// System API/SEC/API/bds_sec_saveSecret
/// This API function is used to store a 16 byte secret key for a specific security access level.
///
///=======
/// Remarks:
///=======
///
///   + The secret keys are stored in an encrypted flash section of the Hardware Security Module (HSM) and cannot be read out.
///   + This asynchronous function must be called several times until the result is available.
///   + If there is no HSM access conflict with another instance, the completion of this function (execution within a loop) takes
///	   + about 1250us (microseconds) with a new secret key and
///	   + about 350us (microseconds) with the same secret key as already stored.
///   + This function will be rejected if another asynchronous security function was already started for this instance.
///
///----------
/// FFI:
///----------
///This API can be used in trusted partitions only. See Freedom from Interference (FFI) concept for more details.
///
///----------
/// Attention:
///----------
///
///   + This function writes the secret key physically into the HSM flash. Therefore this function should not be called cyclically.
///   + Do not interrupt this function by power off to prevent corrupted secret keys.
///
///==================================================================		  			===================================================================================================
///Return value    								  									Description
///==================================================================		  			===================================================================================================
///16#0000: BDS_SEC_ERR_NO_ERROR_DU16													Function was executed without errors. The provided secret key was stored in HSM.
///16#0001: BDS_SEC_ERR_PARAM1_ERROR_DU16												Invalid instance number. 
///16#0002: BDS_SEC_ERR_PARAM2_ERROR_DU16												Invalid access level.
///16#0003: BDS_SEC_ERR_PARAM3_ERROR_DU16												Invalid secret key pointer. Pointer is equal to zero.
///16#0010: BDS_SEC_ERR_REQUEST_PENDING_DU16											This asynchronous function was not yet completed and must be called again with the same parameter values. Several function calls may be required in particular if another security manager instance is also running.
///16#0020:BDS_SEC_ERR_INVALID_SEQUENCE_DU16											This function was called although another asynchronous security function was not yet completed. The other asynchronous function that has already been started must be called again and must be completed before this function can be started.
///16#0033: BDS_SEC_ERR_OPEN_SESSION_FAILED_DU16										Security session could not be opened for this function.Possible reason could be that the HSM is not running. 
///16#0035: BDS_SEC_ERR_CLOSE_SESSION_FAILED_DU16										Security session could not be closed for this function. 
///16#0038: BDS_SEC_ERR_SET_PASSWORD_FAILED_DU16										The internal storage of the secret key failed. To terminate the function, it must be called again.
///
///==================================================================		   			===================================================================================================
///
///For Access levels, Refer the below table & provide the value,
///
///==================================================================		  			===================================================================================================
///Access Level Variable   								  							Value
///==================================================================		  			===================================================================================================
///BDS_SEC_ACC_LEVEL_0_E																0
///BDS_SEC_ACC_LEVEL_1_E																1
///BDS_SEC_ACC_LEVEL_2_E																2
///BDS_SEC_ACC_LEVEL_3_E																3
///BDS_SEC_ACC_LEVEL_4_E																4
///BDS_SEC_ACC_LEVEL_5_E																5
///BDS_SEC_ACC_LEVEL_6_E																6
///BDS_SEC_ACC_LEVEL_7_E																7
///BDS_SEC_ACC_LEVEL_8_E																8
///BDS_SEC_ACC_LEVEL_9_E																9
///BDS_SEC_ACC_LEVEL_10_E																10
///BDS_SEC_ACC_LEVEL_11_E																11
///BDS_SEC_ACC_LEVEL_12_E																12
///BDS_SEC_ACC_LEVEL_13_E																13
///BDS_SEC_ACC_LEVEL_14_E																14
///BDS_SEC_ACC_LEVEL_15_E																15
///BDS_SEC_ACC_LEVEL_16_E																16
///BDS_SEC_ACC_LEVEL_17_E																17
///BDS_SEC_ACC_LEVEL_18_E																18
///BDS_SEC_ACC_LEVEL_19_E																19
///BDS_SEC_ACC_LEVEL_20_E																20
///
///==================================================================		   			===================================================================================================
///
///=======
///Code Example:
///=======
///============================================================================
///
///PROGRAM appl_Task_1
///
///  VAR
///	return_u16 : UINT;
///
///	secKey_au8 : STRING(16);
///	
///  END_VAR
///  
///  (*check for request to store a new secret key*)
///
/// secKey_au8 :=  'MyNewKey' 
///
///result_u16 := bds_sec_saveSecret(bds_diag_inst_te.BDS_SEC_ASW_INST_NAME_1_E, 1, ADR(secKey_au8));
///
///============================================================================
///
{attribute 'external_name' := 'cmp_rts_bds_sec_saveSecret'}
FUNCTION bds_sec_saveSecret : UINT
VAR_INPUT
	///Instance number. pointer to |bds_diag_inst_te|
	diagInst_e: bds_diag_inst_te;
	///Pointer to a variable which must be provided(Refer access level table). The current level will be copied to this variable. 
	level_e: USINT;
	///Pointer to a 16 byte buffer which must be provided by the application and which must contain the new secret key.
	secrKey_pau8: POINTER TO USINT;
END_VAR

END_FUNCTION

// System API/SEC/API/bds_sec_scrambleRexrothSecretsPerm
///This API function is used to scramble all internally stored Rexroth secret keys.
///
///=======
/// Remarks:
///=======
///
///   + This asynchronous function must be called several times until the final result is available.
///   + The completion of this function (execution within a loop) takes about 5,3ms if there is no HSM access conflict with another instance.
///   + This function will be rejected if another asynchronous security function was already started for this instance.
///
///----------
/// FFI:
///----------
///This API can be used in trusted partitions only. See Freedom from Interference (FFI) concept for more details.
///
///----------
/// Attention:
///----------
///
///This function cannot be undone! After the execution of this function the corresponding Rexroth access levels can not be activated any more. This excludes Rexroth personnel from diagnosis information that might be required in case of field service or field claims irrevocably. 
///   
///----------
/// Info:
///----------
///
///This function writes the secret keys physically into the HSM flash. Therefore this function should not be called cyclically.
///   
///==================================================================		  			===================================================================================================
///Return value    								  									Description
///==================================================================		  			===================================================================================================
///16#0000: BDS_SEC_ERR_NO_ERROR_DU16													Function was executed without errors
///16#0010: BDS_SEC_ERR_REQUEST_PENDING_DU16											This asynchronous function was not yet completed and must be called again with the same parameter values. Several function calls may be required in particular if another security manager instance is also running.
///16#0020: BDS_SEC_ERR_INVALID_SEQUENCE_DU16											This function was called although another asynchronous security function was not yet completed. The other asynchronous function that has already been started must be called again and must be completed before this function can be started.
///16#0033: BDS_SEC_ERR_OPEN_SESSION_FAILED_DU16										Security session could not be opened for this function.Possible reason could be that the HSM is not running. 
///16#0034: BDS_SEC_ERR_GENERATE_RANDOM_FAILED_DU16										The process to generate the random has been failed.  To terminate the function, it must be called again.
///16#0035: BDS_SEC_ERR_CLOSE_SESSION_FAILED_DU16										Security session could not be closed for this function. 
///16#0038: BDS_SEC_ERR_SET_PASSWORD_FAILED_DU16										The internal storage of the secret key failed. To terminate the function, it must be called again.
///
///==================================================================		   			===================================================================================================
///
///
///=======
///Code Example:
///=======
///============================================================================
///
///PROGRAM appl_Task_1
///
///  VAR
///	
///  END_VAR
///  
///  (*check if Rexroth access levels shall be scrambled & call the API*)
///  
///result_u16 := bds_sec_scrambleRexrothSecretsPerm();
///
///============================================================================
///
{attribute 'external_name' := 'cmp_rts_bds_sec_scrambleRexrothSecretsPerm'}
FUNCTION bds_sec_scrambleRexrothSecretsPerm : UINT

END_FUNCTION

// System API/SYS/API/bds_sys_ait
///This function gets the temperature of the printed circuit board (PCB)
///
///=======
/// Remarks:
///=======
///    + The voltage of the NTC thermistor located on the PCB is transferred into temperature between -40..150°C.
///    + The resolution is 1°C .
///    + The |GVL_sys| is given for usage of defines.
///    + Import the bds_rts_ec.xml to use the enums. (Refer example below).
///
///----------
/// FFI:
///----------
///This API can be used in trusted partitions only. See Freedom from Interference (FFI) concept for more details.
///
///==================================================================		  			===================================================================================================
///Return value    								  									Description
///==================================================================		  			===================================================================================================
///16#00																				No error.
///16#01																				A parameter is invalid.
///16#02																				Function call was erroneous.
///
///==================================================================		   			===================================================================================================
///
///=======
///Code Example:
///=======
///============================================================================
///
///PROGRAM appl_10ms_task
///
///VAR
///	tsg1_value_s16: INT := 16#00;
///END_VAR
///
///(* get a temperature 1 of high temperature of hardware*)
///
///bds_sys_ait(bds_sys_ait_signal_te.TSGI1, ADR(tsg1_value_s16));
///
///============================================================================
{attribute 'external_name' := 'cmp_rts_bds_sys_ait'}
FUNCTION bds_sys_ait : USINT
VAR_INPUT
	///The assigned signal name of the input.
	signal_e: UINT;
	///Storage address of the value.
	///
	///Range:
	///-40..150 [°C]
	value_ps16: POINTER TO INT;
END_VAR

END_FUNCTION

// System API/SYS/API/bds_sys_aiv
///This function gets the voltage of the analog system input.
///
///=======
/// Remarks:
///=======
///    + Enable the access to all system voltages [mV].
///    + The |GVL_sys| is given for usage of defines.
///    + Import the bds_rts_ec.xml to use the enums. (Refer example below).
///
///----------
/// FFI:
///----------
///This API can be used in trusted partitions only. See Freedom from Interference (FFI) concept for more details.
///	
///==================================================================		  			===================================================================================================
///Return value    								  									Description
///==================================================================		  			===================================================================================================
///16#00																				No error.
///16#01																				A parameter is invalid.
///16#02																				Function call was erroneous.
///
///==================================================================		   			===================================================================================================
///
///=======
///Code Example:
///=======
///============================================================================
///
///PROGRAM appl_10ms_task
///
///VAR
///
///	state_VSS4_u16: UINT := 16#00;
///
///END_VAR
///
///
///(* get a sensor supply voltage *)
///
///bds_sys_aiv(bds_sys_aiv_signal_te.VSS4V10, ADR(state_VSS4_u16));
///
///
///============================================================================
{attribute 'external_name' := 'cmp_rts_bds_sys_aiv'}
FUNCTION bds_sys_aiv : USINT
VAR_INPUT
	///The signal name of the input.
	signal_e: UINT;
	///Storage address of the value.
	///
	///Range:
	///0..40000 [mV]
	value_pu16: POINTER TO UINT;
END_VAR

END_FUNCTION

// System API/SYS/API/bds_sys_cancelAltWakeup
///This function transitions the ECU operating state from RUN to POSTRUN, when the system wakeup reason is not T15. For different methods of ECU wakeup mechanisms please refer page Wakeup.
///
///=======
/// Remarks:
///=======
///    + This function has to be called when the ECU is in RUN state. 
///    + This is most suitable for applications where T15 is not used to switch the ECU OFF.
///    + Wakeup source information can be identified using the BSW API |bds_sys_getResetInfo|.
///    + BSW API |bds_sys_releasePostRunProlong| is used to transition the ECU operating state from POSTRUN to SHUTDOWN.
///    + The |GVL_sys| is given for usage of defines.
///	
///----------
/// FFI:
///----------
///This API can be used in trusted partitions only. See Freedom from Interference (FFI) concept for more details.
///
///----------
/// NOTICE:
///----------
///    + This function has no effect when ECU wakeup has occurred by T15.
///	
///==================================================================		  			===================================================================================================
///Return value    								  									Description
///==================================================================		  			===================================================================================================
///0																					ECU Operating state has moved from RUN to POSTRUN.
///1																					T15 (Ignition pin) is ON.x
///																					    + Note: This return value appears also when ECU woke up by CAN and then T15 turns ON, before this function is called. So, after this, to transition the ECU to POSTRUN state T15 should be turned OFF.
///2																					ECU is already in POSTRUN state.
///
///==================================================================		   			===================================================================================================
///
///=======
///Code Example:
///=======
///============================================================================
///
///PROGRAM PRG
///
///VAR
///
///	return_u8 : USINT;
///
/// flag_u8 :USINT;
///
///END_VAR
///
///IF(0 = flag_u8) THEN
///
/// bds_sys_requestPostRunProlong(); (* request for prolong in POSTRUN*)
///
///	return_u8 := bds_sys_cancelAltWakeup(); (*forces system state to go to POSTRUN*)
///
/// bds_sys_releasePostrunProlong(); (*transitions system state from POSTRUN to SHUTDOWN*)
///
/// flag_u8:=1;
///
///END_IF
///
///============================================================================
{attribute 'external_name' := 'cmp_rts_bds_sys_cancelAltWakeup'}
FUNCTION bds_sys_cancelAltWakeup : USINT

END_FUNCTION

// System API/SYS/API/bds_sys_getResetInfo
///This function can be used in order to get information about reset of ECU.
///
///=======
/// Remarks:
///=======
///    + This function should be used in case of reset problems. The Rexroth service needs this info for solving the problem.
///    + The reset information will only be cleared after power on.
///    + The Reset IDs & Reset Group IDs can be found in "rba_Reset_Cfg.h" header file. All the Reset group IDs are listed down under enum variable "rba_Reset_Grp_ten" and all the reset IDs are listed down under enum variable "rba_Reset_Id_ten".
///    + The |GVL_sys| is given for usage of defines.
///
///----------
/// FFI:
///----------
///This API can be used in trusted partitions . For untrusted partitions use |bds_sys_getResetInfo_ffi|. See Freedom from Interference (FFI) concept for more details.
///
///==================================================================		  			===================================================================================================
///Return value    								  									Description
///==================================================================		  			===================================================================================================
///16#0000																				No error. 
///16#0001																				Function called with null pointer.
///16#25																				FFI API access error.
///
///==================================================================		   			===================================================================================================
///=======
///Code Example:
///=======
///============================================================================
///
///PROGRAM appl_10ms_task
///
///VAR
///
///	reset_info : bds_ResetInfo_ts;
///	
///	return_u8 : UINT;
///
///END_VAR
///
///return_u8 := bds_sys_getResetInfo(ADR(reset_info)); (*reads the reset information of ECU*)
///
///============================================================================
{attribute 'external_name' := 'cmp_rts_bds_sys_getResetInfo'}
FUNCTION bds_sys_getResetInfo : UINT
VAR_INPUT
	///Pointer to |bds_ResetInfo_ts|
	resetinfo_ps: POINTER TO bds_ResetInfo_ts;
END_VAR

END_FUNCTION

// System API/SYS/FFI_API/bds_sys_getResetInfo_ffi
{attribute 'external_name' := 'cmp_rts_bds_sys_getResetInfo_ffi'}
FUNCTION bds_sys_getResetInfo_ffi : UINT
VAR_INPUT
	///Pointer to |bds_ResetInfo_ts|
	resetinfo_ps: POINTER TO bds_ResetInfo_ts;
END_VAR

END_FUNCTION

// System API/SYS/API/bds_sys_releasePostRunProlong
///This function terminates prolonging of  POSTRUN state and enters to SHUTDOWN state.     
///=======
/// Remarks:
///=======
///    + By calling this function, POSTRUN is terminated, if system is in POSTRUN state and enters to SHUTDOWN phase. 
///    + After calling |bds_sys_requestPostRunProlong| and after completion of tasks in POSTRUN this function must be called. If not, exit from POSTRUN is only through timeout.
///    + The |GVL_sys| is given for usage of defines.
///	
///----------
/// FFI:
///----------
///This API can be used in trusted partitions only. See Freedom from Interference (FFI) concept for more details.
///
///==================================================================		  			===================================================================================================
///Return value    								  									Description
///==================================================================		  			===================================================================================================
///None																				None
///
///==================================================================		   			===================================================================================================
///
///
///=======
///Code Example:
///=======
///============================================================================
///
///PROGRAM appl_1ms_task
///
///VAR
///
///END_VAR
///
///bds_sys_releasePostRunProlong();  (* release of prolong in postrun *)
///
///============================================================================
{attribute 'external_name' := 'cmp_rts_bds_sys_releasePostRunProlong'}
FUNCTION bds_sys_releasePostRunProlong : BOOL

END_FUNCTION

// System API/SYS/API/bds_sys_requestPostRunProlong
///This function enables a prolonging cyclic tasks in POSTRUN.    
///=======
/// Remarks:
///=======
///    + This function can be called in initialization or RUN state of system.
///    + After calling this function, termination from POSTRUN state is possible only by calling |bds_sys_releasePostRunProlong| or Timeout set for POSTRUN prolong.  
///    + The Maximum Post Run timeout allowed is 24hours / 86400 sec. The actual Post Run timeout is configured in easyConfig.In order to shorten the Post Run timeout  the  API |bds_sys_releasePostRunProlong| shall be used.
///    + Without calling this function, No cyclic tasks are in POSTRUN. Only shutdown functions will be executed after Ignition(T15) goes OFF.
///    + The |GVL_sys| is given for usage of defines.
///	
///----------
/// FFI:
///----------
///This API can be used in trusted partitions only. See Freedom from Interference (FFI) concept for more details.
///
///---------
///  NOTICE:
///---------
///Don't forget to call  |bds_sys_releasePostRunProlong|, after enabling cyclic tasks POSTRUN.
///	
///==================================================================		  			===================================================================================================
///Return value    								  									Description
///==================================================================		  			===================================================================================================
///None																				None
///
///==================================================================		   			===================================================================================================
///
///
///=======
///Code Example:
///=======
///============================================================================
///
///PROGRAM appl_1ms_task
///
///VAR
///
///END_VAR
///
///bds_sys_requestPostRunProlong();  (* request for prolong in postrun *)
///
///============================================================================
{attribute 'external_name' := 'cmp_rts_bds_sys_requestPostRunProlong'}
FUNCTION bds_sys_requestPostRunProlong : BOOL

END_FUNCTION

// System API/SYS/API/bds_sys_di
///This function gets the state of a digital system input.
///
///=======
/// Remarks:
///=======
///    + Enable the access to all digital signals.
///    + The |GVL_sys| is given for usage of defines.
///    + Import the bds_rts_ec.xml to use the enums. (Refer example below).
///
///----------
/// FFI:
///----------
///This API can be used in trusted partitions only. See Freedom from Interference (FFI) concept for more details.
///
///==================================================================		  			===================================================================================================
///Return value    								  									Description
///==================================================================		  			===================================================================================================
///16#00																				No error.
///16#01																				A parameter is invalid.
///16#02																				Function call was erroneous.
///
///==================================================================		   			===================================================================================================
///
///=======
///Code Example:
///=======
///============================================================================
///
///PROGRAM appl_10ms_task
///
///VAR
///
///	state_u8: USINT := 16#00;
///
///END_VAR
///
///(* get a state of the inhibit signal *)
///
///bds_sys_di(bds_sys_di_signal_te.ST_INH, ADR(state_u8));
///
///============================================================================
{attribute 'external_name' := 'cmp_rts_bds_sys_di'}
FUNCTION bds_sys_di : USINT
VAR_INPUT
	///The assigned signal name of the input.
	signal_e: UINT;
	///Storage address of the state.
	///
	///States:
	///    + 0 : OFF
	///    + 1 : ON
	state_pu8: POINTER TO USINT;
END_VAR

END_FUNCTION

// System API/SYS/API/bds_sys_getAge
///This function reads the operating time counter of the ECU in minutes.
///
///=======
/// Remarks:
///=======
///    + The counter is incremented by 1 for each minute and saved in non-volatile memory for every 30 minutes.
///    + The operating time counter cannot be reset.
///    + The operating time counter records the total operating time of the device in minutes.
///    + The system time of controller since last reset can be determined using the functions |bds_sys_getTime|.
///    + The |GVL_sys| is given for usage of defines.
///	
///----------
/// FFI:
///----------
///This API can be used in trusted partitions . For untrusted partitions use |bds_sys_getAge_ffi|. See Freedom from Interference (FFI) concept for more details.
///
///----------
/// NOTICE:
///----------
///    + Operating time is saved in case of ignition off event
///    + Operation time is not saved, if ECU power supply is switched off .
///
///==================================================================		  			===================================================================================================
///Return value    								  									Description
///==================================================================		  			===================================================================================================
///Value																				Total operating time of the ECU in minutes
///16#00: BDS_SYS_FFI_ACCESS_ERROR_GETVALUE_DU32										FFI API access error.
///
///==================================================================		   			===================================================================================================
///
///=======
///Code Example:
///=======
///============================================================================
///
///PROGRAM appl_10ms_task
///
///VAR
///
///	operating_hours_u32: UDINT := 16#00;
///
///END_VAR
///
///operating_hours_u32 := bds_sys_getAge(); (* returns Total operating hours of the ECU in minutes *)
///
///============================================================================
{attribute 'external_name' := 'cmp_rts_bds_sys_getAge'}
FUNCTION bds_sys_getAge : UDINT

END_FUNCTION

// System API/SYS/API/bds_sys_getTime
///This function reads the system time of controller since last reset.
///=======
/// Remarks:
///=======
///    + The system time starts at 0 again every time the system is switched on. 
///    + Return value is 64 bit value (counter width).
///    + In order to detect a counter overrun, for long operating times, the operating time counter must also be evaluated using the function |bds_sys_getAge|. 
///    + The |GVL_sys| is given for usage of defines.
///
///----------
/// FFI:
///----------
///This API can be used in trusted partitions . For untrusted partitions use |bds_sys_getTime_ffi|. See Freedom from Interference (FFI) concept for more details.
///
///==================================================================		  			===================================================================================================
///Return value    								  									Description
///==================================================================		  			===================================================================================================
///Value																				System time in microseconds [us].
///16#00: BDS_SYS_FFI_ACCESS_ERROR_GETVALUE_DU64										FFI API access error.
///
///==================================================================		   			===================================================================================================
///
///
///=======
///Code Example:
///=======
///============================================================================
///
///PROGRAM appl_10ms_task
///
///VAR
///
///	operating_time : ULINT := 16#00;
///
///END_VAR
///
///operating_time := bds_sys_getTime();  (* returns Operating time in microseconds since last reset *)
///
///============================================================================
{attribute 'external_name' := 'cmp_rts_bds_sys_getTime'}
FUNCTION bds_sys_getTime : ULINT

END_FUNCTION

// System API/SYS/FFI_API/bds_sys_getTime_ffi
{attribute 'external_name' := 'cmp_rts_bds_sys_getTime_ffi'}
FUNCTION bds_sys_getTime_ffi : ULINT

END_FUNCTION

// System API/SYS/FFI_API/bds_sys_getAge_ffi
{attribute 'external_name' := 'cmp_rts_bds_sys_getAge_ffi'}
FUNCTION bds_sys_getAge_ffi : UDINT

END_FUNCTION

// System API/SYS/API/bds_sys_getCoreLoad
///This function will provide core load for a specified core in percentage.
///
///=======
/// Remarks:
///=======
///    + Current Cycle Max Load and Life Cycle Max Load is also provided for a specified core in percentage.
///    + Core load is the load in the elapsed time frame.
///    + Core load,Current Cycle Max Load and Life Cycle Max Load is in percentage with resolution of 0.01%.
///    + All the application tasks present in Core 1.
///    + The |GVL_sys| is given for usage of defines.
///	
///----------
/// FFI:
///----------
///This API can be used in trusted partitions . For untrusted partitions use |bds_sys_getCoreLoad_ffi|. See Freedom from Interference (FFI) concept for more details.
///
///----------
/// NOTICE:
///----------
///For load on CPU check the load on Core1.
///
///==================================================================		  			===================================================================================================
///Return value    								  									Description
///==================================================================		  			===================================================================================================
///16#00																				No Errors.
///16#01																				Wrong Core ID.
///16#02																				Invalid Pointer.
///16#25																				FFI API access error.
///
///==================================================================		   			===================================================================================================
///=======
///Code Example:
///=======
///============================================================================
///
///PROGRAM appl_10ms_task
///
///VAR
///
///	coreID_e : bds_sys_coreid_te;
///
///	core_load  : bds_sys_coreload_info_ts;
///
///	status_u8 : USINT;
///
///END_VAR
///
///status_u8 := bds_sys_getCoreLoad(coreID_e,ADR(core_load)); (*Function for getting the Core load*)
///
///============================================================================
{attribute 'external_name' := 'cmp_rts_bds_sys_getCoreLoad'}
FUNCTION bds_sys_getCoreLoad : USINT
VAR_INPUT
	///Logical ID of the Core
	coreID_e: bds_sys_coreid_te;
	///Storage address for the core load.
	///	
	///Pointer to the |bds_sys_coreload_info_ts|
	core_load_ps: POINTER TO bds_sys_coreload_info_ts;
END_VAR

END_FUNCTION

// System API/SYS/FFI_API/bds_sys_getCoreLoad_ffi
{attribute 'external_name' := 'cmp_rts_bds_sys_getCoreLoad_ffi'}
FUNCTION bds_sys_getCoreLoad_ffi : USINT
VAR_INPUT
	///Logical ID of the Core
	coreID_e: bds_sys_coreid_te;
	///Storage address for the core load.
	///	
	///Pointer to the |bds_sys_coreload_info_ts|
	core_load_ps: POINTER TO bds_sys_coreload_info_ts;
END_VAR

END_FUNCTION

// System API/SYS/API/bds_sys_getEcuInfo
///This function gets information of ECU from System Memory Page.
///
///=======
/// Remarks:
///=======
///    + The |GVL_sys| is given for usage of defines.
///	
///----------
/// FFI:
///----------
///This API can be used in trusted partitions . For untrusted partitions use |bds_sys_getEcuInfo_ffi|. See Freedom from Interference (FFI) concept for more details.
///
///==================================================================		  			===================================================================================================
///Return value    								  									Description
///==================================================================		  			===================================================================================================
///16#0000																				No error.
///16#0001																				No correct ECU information.
///16#0002																				Function is called with NULL pointer.
///16#25																				FFI API access error.
///
///==================================================================		   			===================================================================================================
///
///=======
///Code Example:
///=======
///============================================================================
///
///PROGRAM appl_100ms_task
///
///VAR
///
///	EcuInfo_s: bds_EcuInfo_ts;
///
///	return_u16: UINT := 16#00; 
///
///END_VAR
///
///return_u16 := bds_sys_getEcuInfo(ADR(EcuInfo_s));
///
///
///============================================================================
{attribute 'external_name' := 'cmp_rts_bds_sys_getEcuInfo'}
FUNCTION bds_sys_getEcuInfo : UINT
VAR_INPUT
	///Pointer to |bds_EcuInfo_ts|
	EcuInfo_ps: POINTER TO bds_EcuInfo_ts;
END_VAR

END_FUNCTION

// System API/SYS/FFI_API/bds_sys_getEcuInfo_ffi
{attribute 'external_name' := 'cmp_rts_bds_sys_getEcuInfo_ffi'}
FUNCTION bds_sys_getEcuInfo_ffi : UINT
VAR_INPUT
	///Pointer to |bds_EcuInfo_ts|
	EcuInfo_ps: POINTER TO bds_EcuInfo_ts;
END_VAR

END_FUNCTION

// System API/SYS/API/bds_sys_getStates
///This function gets the current and previous state of system. 
///
///=======
/// Remarks:
///=======
///    + This function should be used in case of reset problems. The Rexroth service needs this info for solving the problem.
///    + The reset information will only be cleared after power on.
///    + The Reset IDs & Reset Group IDs can be found in "rba_Reset_Cfg.h" header file. All the Reset group IDs are listed down under enum variable "rba_Reset_Grp_ten" and all the reset IDs are listed down under enum variable "rba_Reset_Id_ten".
///    + The |GVL_sys| is given for usage of defines.
///
///----------
/// FFI:
///----------
///This API can be used in trusted partitions . For untrusted partitions use |bds_sys_getStates_ffi|. See Freedom from Interference (FFI) concept for more details.
///	
///---------
///  NOTICE:
///---------
///During power on initialization current and previous states are same.
///
///==================================================================		  			===================================================================================================
///Return value    								  									Description
///==================================================================		  			===================================================================================================
///16#00																				No error.
///16#01																				A parameter is invalid.
///16#25																				FFI API access error.
///
///==================================================================		   			===================================================================================================
///
///=======
///Code Example:
///=======
///============================================================================
///
///PROGRAM appl_10ms_task
///
///VAR
///
///	states_s: bds_sys_states_ts;
///
///	return_u8: USINT := 16#00;
///
///END_VAR
///
///return_u8 := bds_sys_getStates(ADR(states_s));  (* read current and previous states of system. *)
///
///============================================================================
{attribute 'external_name' := 'cmp_rts_bds_sys_getStates'}
FUNCTION bds_sys_getStates : USINT
VAR_INPUT
	///Storage address for the systems states.
	///	
	///The different system states are:
	///
	///    + BDS_SYSSTATE_INIT_E (0)
	///    + BDS_SYSSTATE_RUN_E(1)
	///    + BDS_SYSSTATE_POSTRUN_E(2)
	///    + BDS_SYSSTATE_SHUTDOWN_E(3)
	states_ps: POINTER TO bds_sys_states_ts;
END_VAR

END_FUNCTION

// System API/SYS/FFI_API/bds_sys_getStates_ffi
{attribute 'external_name' := 'cmp_rts_bds_sys_getStates_ffi'}
FUNCTION bds_sys_getStates_ffi : USINT
VAR_INPUT
	///Storage address for the systems states.
	///	
	///The different system states are:
	///
	///    + BDS_SYSSTATE_INIT_E (0)
	///    + BDS_SYSSTATE_RUN_E(1)
	///    + BDS_SYSSTATE_POSTRUN_E(2)
	///    + BDS_SYSSTATE_SHUTDOWN_E(3)
	states_ps: POINTER TO bds_sys_states_ts;
END_VAR

END_FUNCTION

// System API/SYS/API/bds_sys_getT15
///This function gets the state of the terminal input T15 (Ignition).
///
///=======
/// Remarks:
///=======
///    + The state of the terminal input T15 is the debounced signal.
///    + The |GVL_sys| is given for usage of defines.
///
///----------
/// FFI:
///----------
///This API can be used in trusted partitions only. See Freedom from Interference (FFI) concept for more details.
///
///==================================================================		  			===================================================================================================
///Return value    								  									Description
///==================================================================		  			===================================================================================================
///None.																				None.
///
///==================================================================		   			===================================================================================================
///
///=======
///Code Example:
///=======
///============================================================================
///
///PROGRAM appl_10ms_task
///
///VAR
///
///	tT15_u8: USINT := 16#00;
///
///END_VAR
///
///(* get state of T15 *)
///
///bds_sys_getT15(ADR(tT15_u8));
///
///
///============================================================================
{attribute 'external_name' := 'cmp_rts_bds_sys_getT15'}
FUNCTION bds_sys_getT15 : BOOL
VAR_INPUT
	///Storage address of the state.
	///
	///States:
	///    + 0 : OFF
	///    + 1 : ON
	stT15_pu8: POINTER TO USINT;
END_VAR

END_FUNCTION

// System API/SYS/API/bds_sys_getTaskRuntime
///This function will provide task runtime of a specified task in microseconds. 
///
///=======
/// Remarks:
///=======
///    + Task Load consists of Gross Runtime (inclusive of Interrupts) and Net Runtime (exclusive of Interrupts).
///    + All the values of task load are in microseconds.
///    + Number of tasks for which BSW provides the measurement are (1ms,10ms,20ms,40ms,50ms,80ms,100ms).  
///    + The |GVL_sys| is given for usage of defines.
///
///----------
/// FFI:
///----------
///This API can be used in trusted partitions . For untrusted partitions use |bds_sys_getTaskRuntime_ffi|. See Freedom from Interference (FFI) concept for more details.
///
///==================================================================		  			===================================================================================================
///Return value    								  										Description
///==================================================================		  			===================================================================================================
///16#00																				No Error.
///16#01																				Wrong Task ID.
///16#02																				Invalid Pointer.
///16#25																				FFI API access error.
///
///==================================================================		   			===================================================================================================
///=======
///Code Example:
///=======
///============================================================================
///
///PROGRAM appl_10ms_task
///
///VAR
///
///	task_runtime : bds_sys_taskruntime_ts ;
///	
///	return_u8 : UINT;
///
///END_VAR
///
///return_u8 := bds_sys_getTaskRuntime(bds_sys_task_te.Task_20ms_D , ADR(task_runtime)); (*Function for getting task runtime*)
///
///============================================================================
{attribute 'external_name' := 'cmp_rts_bds_sys_getTaskRuntime'}
FUNCTION bds_sys_getTaskRuntime : USINT
VAR_INPUT
	///Task Id for which task load is required
	task_name_e: bds_sys_task_te;
	///Storage address for the Task Load
	///pointer to |bds_sys_getTaskRuntime|
	task_runtime_ps: POINTER TO bds_sys_taskruntime_ts;
END_VAR

END_FUNCTION

// System API/SYS/FFI_API/bds_sys_getTaskRuntime_ffi
{attribute 'external_name' := 'cmp_rts_bds_sys_getTaskRuntime_ffi'}
FUNCTION bds_sys_getTaskRuntime_ffi : USINT
VAR_INPUT
	///Task Id for which task load is required
	task_name_e: bds_sys_task_te;
	///Storage address for the Task Load
	///pointer to |bds_sys_getTaskRuntime|
	task_runtime_ps: POINTER TO bds_sys_taskruntime_ts;
END_VAR

END_FUNCTION

// System API/SYS/API/bds_sys_getVersion
///This function gets the name and version of software parts (modules).
///=======
/// Remarks:
///=======
///    + The |GVL_sys| is given for usage of defines.
///
///----------
/// FFI:
///----------
///This API can be used in trusted partitions . For untrusted partitions use |bds_sys_getVersion_ffi|. See Freedom from Interference (FFI) concept for more details.
///
///==================================================================		  			===================================================================================================
///Return value    								  									Description
///==================================================================		  			===================================================================================================
///BDS_SYSGETVERSION_OK_DU16 (16#00)													 No error.
///BDS_SYSGETVERSION_BUFLEN_UNDERSIZE_DU16 (16#01)										The given buffer (buf_pau8 / bufLen_u16) is to small to be able to receive the complete version data. The data was truncated to the given buffer length.
///BDS_SYSGETVERSION_SW_PART_INVALID_DU16 (16#02)										Invalid software part.
///BDS_SYSGETVERSION_SW_INFO_NOT_FOUND_DU16 (16#03)									Software part info not found.
///BDS_SYSGETVERSION_BUF_INVALID_DU16 (16#04)I											nvalid pointer for data buffer.
///BDS_SYSGETVERSION_COPIEDBYTES_INVALID_DU16 (16#05)									Invalid pointer for number of copied bytes.
///16#25																				FFI API access error.
///
///
///==================================================================		   			===================================================================================================
///
///
///=======
///Code Example:
///=======
///============================================================================
///
///VAR_GLOBAL CONSTANT
///
///	myBufLen_DU8: USINT := 64;
///
///END_VAR
///
/// 
///
///PROGRAM appl_100ms_task
///
///VAR
///
///	myBufData_au8: ARRAY[1..myBufLen_DU8] OF USINT;
///
///	copiedBytes_u16: UINT := 16#00;
///
///	retVal_u16: UINT := 16#00;
///
///END_VAR
///
///(* get application software name *)
///
///retVal_u16 := bds_sys_getVersion(BDS_VERSION_SW_PART_APPL_DU8, ADR(myBufData_au8), myBufLen_DU8, ADR(copiedBytes_u16));
///
/// 
///
///IF BDS_SYSGETVERSION_OK_DU16 = retVal_u16 THEN
///
///  (* the first copiedBytes_u16 bytes in myBufData_au8[] can be evaluated here *)
///
///END_IF
///
///
///============================================================================
{attribute 'external_name' := 'cmp_rts_bds_sys_getVersion'}
FUNCTION bds_sys_getVersion : UINT
VAR_INPUT
	///Selection of the software part (module):
	///    + BDS_VERSION_SW_PART_APPL_DU8  (Application software name from bds_sysInit())    
	///    + BDS_VERSION_SW_PART_SB_DU8  (Bootcontrol start up module)         
	///    + BDS_VERSION_SW_PART_CB_DU8  (Customer boot loader module)         
	///    + BDS_VERSION_SW_PART_BSW_NAME_DU8  (Name of BSW)  
	///    + BDS_VERSION_SW_PART_BSW_VERSION_DU8  (Version of BSW)
	///    + BDS_VERSION_SW_PART_EC_PROJECT_DU8  (EasyConfig project name)
	swPart_u8: USINT;
	///Pointer to buffer which will be used to return version data. The number of bytes which can be written by API is specified in parameter bufLen_u16.
	buf_pau8: POINTER TO USINT;
	///Length of the buffer in bytes specified with buf_pau8.
	bufLen_u16: UINT;
	///Pointer to a variable which will be used to return the number of valid data in buffer specified by buf_pu8.
	copiedBytes_pu16: POINTER TO UINT;
END_VAR

END_FUNCTION

// System API/SYS/FFI_API/bds_sys_getVersion_ffi
{attribute 'external_name' := 'cmp_rts_bds_sys_getVersion_ffi'}
FUNCTION bds_sys_getVersion_ffi : UINT
VAR_INPUT
	///Selection of the software part (module):
	///    + BDS_VERSION_SW_PART_APPL_DU8  (Application software name from bds_sysInit())    
	///    + BDS_VERSION_SW_PART_SB_DU8  (Bootcontrol start up module)         
	///    + BDS_VERSION_SW_PART_CB_DU8  (Customer boot loader module)         
	///    + BDS_VERSION_SW_PART_BSW_NAME_DU8  (Name of BSW)  
	///    + BDS_VERSION_SW_PART_BSW_VERSION_DU8  (Version of BSW)
	///    + BDS_VERSION_SW_PART_EC_PROJECT_DU8  (EasyConfig project name)
	swPart_u8: USINT;
	///Pointer to buffer which will be used to return version data. The number of bytes which can be written by API is specified in parameter bufLen_u16.
	buf_pau8: POINTER TO USINT;
	///Length of the buffer in bytes specified with buf_pau8.
	bufLen_u16: UINT;
	///Pointer to a variable which will be used to return the number of valid data in buffer specified by buf_pu8.
	copiedBytes_pu16: POINTER TO UINT;
END_VAR

END_FUNCTION

// System API/SYS/API/bds_sys_getVSS
///This function gets the state of the sensor supply voltage.
///=======
/// Remarks:
///=======
///    + For the sensor supplies VSS1 and VSS2 only the states can be read, there is no possibility to get the sensor voltages.
///    + For the other sensor supplies the function cannot be used, but therefore the sensor voltage can be read with |bds_sys_aiv|.
///    + For the further information regarding diagnostic and the recovery see Cyclic monitoring checks.
///    + The |GVL_sys| is given for usage of defines.
///    + Import the bds_rts_ec.xml to use the enums. (Refer example below).
///
///----------
/// FFI:
///----------
///This API can be used in trusted partitions only. See Freedom from Interference (FFI) concept for more details.
///
///==================================================================		  			===================================================================================================
///Return value    								  									Description
///==================================================================		  			===================================================================================================
///16#00																				No error.
///16#01																				A parameter is invalid.
///16#02																				Function call was erroneous.
///
///==================================================================		   			===================================================================================================
///
///
///=======
///Code Example:
///=======
///============================================================================
///
///PROGRAM appl_10ms_task
///
///VAR
///
///	stVSS1_u8: USINT := 16#00;
///
///END_VAR
/// 
///
///(* get state of VSS1 *)
///
///bds_sys_getVSS(bds_sys_vss_signal_te.VSS1, ADR(stVSS1_u8));
///
///
///============================================================================
{attribute 'external_name' := 'cmp_rts_bds_sys_getVSS'}
FUNCTION bds_sys_getVSS : USINT
VAR_INPUT
	///The assigned signal name.
	///
	///Only VSS1 and VSS2 are allowed.
	signal_e: UINT;
	///Storage address of the state.
	///	
	///States:
	///    + 0 : OFF
	///    + 1 : ON
	state_pu8: POINTER TO USINT;
END_VAR

END_FUNCTION

// System API/SYS/API/BDS_SYS_GET_LOCK_COMMON
///Mark an entry into an user critical section. That means nested interrupts are not possible and access to user global variable is safe.     
///
///=======
/// Attention:
///=======
///    + Function |BDS_SYS_RELEASE_LOCK_COMMON| has to be used in order to leave a critical section which is entered.
///    + Stay in a critical section only for a short time! Otherwise e.g. CAN messages can be lost. 
///    + A critical section has to be completed in a function. (That means it is not possible to enter into a critical section in one function and to leave this critical section in another function.)
///
///----------
/// FFI:
///----------
///This API can be used in trusted partitions only. See Freedom from Interference (FFI) concept for more details.
///
///==================================================================		  			===================================================================================================
///Return value    								  									Description
///==================================================================		  			===================================================================================================
///None																				None
///
///==================================================================		   			===================================================================================================
///
///=======
///Code Example:
///=======
///============================================================================
///
///PROGRAM appl
///
///  (*Nested interrupts are possible.*)
/// 
///  BDS_SYS_GET_LOCK_COMMON();
/// 
///  (*No nested interrupts.*)
///  
///  BDS_SYS_RELEASE_LOCK_COMMON();
///  (*Nested interrupts are possible.*)
///
///============================================================================
///
{attribute 'external_name' := 'cmp_rts_BDS_SYS_GET_LOCK_COMMON'}
FUNCTION BDS_SYS_GET_LOCK_COMMON : BOOL

END_FUNCTION

// System API/SYS/API/BDS_SYS_RELEASE_LOCK_COMMON
///Leave an user critical section.     
///
///=======
/// Attention:
///=======
///    + Function |BDS_SYS_GET_LOCK_COMMON| has to be used in order to enter into a critical section.
///    + A critical section has to be completed in a function. (That means it is not possible to enter into a critical section in one function and to leave this critical section in another function.)
///	
///----------
/// FFI:
///----------
///This API can be used in trusted partitions only. See Freedom from Interference (FFI) concept for more details.
///
///==================================================================		  			===================================================================================================
///Return value    								  									Description
///==================================================================		  			===================================================================================================
///None																				None
///
///==================================================================		   			===================================================================================================
///=======
///Code Example:
///=======
///============================================================================
///
///PROGRAM appl
///
///  (*Nested interrupts are possible.*)
/// 
///  BDS_SYS_GET_LOCK_COMMON();
/// 
///  (*No nested interrupts.*)
///  
///  BDS_SYS_RELEASE_LOCK_COMMON();
///  (*Nested interrupts are possible.*)
///
///============================================================================
{attribute 'external_name' := 'cmp_rts_BDS_SYS_RELEASE_LOCK_COMMON'}
FUNCTION BDS_SYS_RELEASE_LOCK_COMMON : BOOL

END_FUNCTION

// System API/SYS/API/bds_sys_memByteCopy
///Memory copy routine, this function will copy the data from one source to another.
///=======
/// Remarks:
///=======
///    + This function must be called to fill the buffer for example in callbacks.
///    + Source and Destination must not be overlapped.
///    + The |GVL_sys| is given for usage of defines.
///
///----------
/// FFI:
///----------
///This API can be used in trusted partitions only. See Freedom from Interference (FFI) concept for more details.
///
///==================================================================		  			===================================================================================================
///Return value    								  									Description
///==================================================================		  			===================================================================================================
///None																				None
///
///==================================================================		   			===================================================================================================
///=======
///Code Example:
///=======
///============================================================================
///
///PROGRAM appl_1ms_task
///
///VAR
///
///	myBufData1_au8: ARRAY[1..3] OF UINT;
///
///	myBufData2_au8: ARRAY[1..3] OF UINT;
///
///	status: BOOL;
///
///END_VAR
///
///myBufData1_au8[1] := 9;
///
///status := bds_sys_memByteCopy(ADR(myBufData1_au8),ADR(myBufData2_au8),3);
///
///
///============================================================================
{attribute 'external_name' := 'cmp_rts_bds_sys_memByteCopy'}
FUNCTION bds_sys_memByteCopy : BOOL
VAR_INPUT
	///Reference of destination variable which needs to be filled. 
	xDest_pu8: POINTER TO USINT;
	///Reference of source variable.
	xSrc_pcu8: POINTER TO USINT;
	///Length of the data bytes which will be copied into buffer.
	numBytes_u32: UDINT;
END_VAR

END_FUNCTION

// System API/SYS/API/bds_sys_resetCoreLoad
///This function will reset the current cycle max load and lifetime cycle max load of all CPU cores.    
///=======
/// Remarks:
///=======
///    + Current cycle max load is set equal to current core load value when the reset operation was performed.
///    + Lifetime cycle max load is set equal to current cycle max load  value when the reset operation was performed.
///    + The |GVL_sys| is given for usage of defines.
///
///	
///----------
/// FFI:
///----------
///This API can be used in trusted partitions only. See Freedom from Interference (FFI) concept for more details.
///
///==================================================================		  			===================================================================================================
///Return value    								  									Description
///==================================================================		  			===================================================================================================
///None																				None
///
///==================================================================		   			===================================================================================================
///=======
///Code Example:
///=======
///============================================================================
///
///PROGRAM appl_1ms_task
///
///VAR
///
///END_VAR
///
///  (*Reset Current Cycle Max Load and LifeTimeCycle max load*)
///
///   bds_sys_resetCoreLoad();
///
///
///============================================================================
///
{attribute 'external_name' := 'cmp_rts_bds_sys_resetCoreLoad'}
FUNCTION bds_sys_resetCoreLoad : BOOL

END_FUNCTION

// System API/SYS/API/bds_sys_resetEcu
///This function resets the ECU.   
///=======
/// Remarks:
///=======
///    + Before this function call bds_sys_resetEcu(), the memory blocks which need to be saved in NVM (NVM general description) should be marked by calling the function |bds_mem_markBlock|. Thus during reset preparation marked memory block is saved into NVM and it can be retrieved after reset. So, it is recommended to call this function with NVMWrite_I = TRUE.
///    + The reset info can be analyzed at the next start up by using the function |bds_sys_getResetInfo|.
///    + The |GVL_sys| is given for usage of defines.
///
///----------
/// FFI:
///----------
///This API can be used in trusted partitions only. See Freedom from Interference (FFI) concept for more details.
///
///==================================================================		  			===================================================================================================
///Return value    								  									Description
///==================================================================		  			===================================================================================================
///None																				None
///
///==================================================================		   			===================================================================================================
///
///
///==================================================================		  			===================================================================================================
///Reset Parameter    								  									Description
///==================================================================		  			===================================================================================================
///Reset Reason  - Reset Group ID														RBA_RESET_GRP_SOFTRESET_E (16#09).
///Reset Reason  - Reset number														RBA_RESET_NUM_ASW (16#304E).
///
///==================================================================		   			===================================================================================================
///
///
///=======
///Code Example:
///=======
///============================================================================
///
///PROGRAM appl_1ms_task
///
///VAR
///
///    Mark_writeval: USINT:=0;
///
///END_VAR
///
///(*Call the markblock API once. Mark the block(eg:3rd block) which has to be written during afterrun cycle in either cyclic task or calling once & assign a value to Mark_writeval*)
///
///bds_mem_markBlock(3,ADR(Mark_writeval),1,1,TRUE);
///
///bds_sys_resetEcu(0x1234, TRUE);
///
///============================================================================
///
{attribute 'external_name' := 'cmp_rts_bds_sys_resetEcu'}
FUNCTION bds_sys_resetEcu : BOOL
VAR_INPUT
	///User defined value which can be used e.g., for Diagnostics
	///
	///    + This user defined value can be retrieved by calling |bds_sys_getResetInfo| function, the output of this function gives out a variable "rbr_UserDefined_u32" which is same as this variable.
	value_u32: UDINT;
	///If the “NVMWrite_l” flag is set to the following values the behaviour is different,
	///    + TRUE   : Function will return and reset will be executed until NVM update is finished.
	///    + FALSE  : Function never return and execute reset immediately.
	NVMWrite_l: BOOL;
END_VAR

END_FUNCTION

// Memory API/NVM/API/bds_mem_markBlock
///This function sets a marker for writing the block data from RAM mirror into corresponding NVM block during next ECU after run.
///
///=======
/// Remarks:
///=======
///
///    + All marked RAM mirrors of the application NVM blocks are automatically written into NVM during after run.
///    + The |GVL_mem| is given for usage of defines.
///
///----------
/// FFI:
///----------
///    + This API can be used in trusted partitions . For untrusted partitions use |bds_mem_markBlock_ffi|. See Freedom from Interference (FFI) concept for more details.
///    + The blocks which can be written using |bds_mem_markBlock_ffi| are mentioned in page NVM block description.
///
///----------
/// NOTICE:
///----------
///    + This function has to called for all these blocks which shall be written into NVM automatically during after run.
///    + If |bds_mem_readBlock| is used after |bds_mem_markBlock| for a particular NVM block, |bds_mem_markBlock| has to be called again for the same NVM block during the same driving cycle before AfterRun.
///
///
///==================================================================		  			===================================================================================================
///Return value    								  									Description
///==================================================================		  			===================================================================================================
///16#0000: BDS_MEM_NO_ERROR_DU16														Reading of block was successfully started.
///16#0001: BDS_MEM_INVALID_BLOCKID_DU16												Invalid Block ID.
///16#0400: BDS_MEM_MARKBLOCK_ERROR_DU16												Read block could not be started e.g. due to actual block status.
///16#0300: BDS_MEM_MARKBLOCK_DATASIZE_INVALID_DU16									Marking the block fails as the data size not fitting into NVM Block
///16#0301: BDS_MEM_MARKBLOCK_DATAPTR_INVALID_DU16										Invalid Data Address
///16#000C: BDS_MEM_FFI_ACCESS_ERROR_DU16												Invalid Access to FFI variant API call.
///
///==================================================================		   			===================================================================================================
///
///=======
///Code Example:
///=======
///============================================================================
///
///PROGRAM markblock
///
///VAR
///
///    Mark_writeval: USINT:=0;
///
///    Readval: USINT:=0;
///
///    ts_mem_mark: UINT;
///
///END_VAR
///
///(*Call the markblock API. Mark the block(eg:78rd block) which has to be written during afterrun cycle in either cyclic task or calling once & assign a value to Mark_writeval*)
///
///ts_mem_mark:=bds_mem_markBlock(78,ADR(Mark_writeval),100,1,TRUE);
///
///(*Switch ignition line off (T15). Wait until ECU is really switched off -> check current (drops to zero). Switch ignition line (T15) on again*)
///
///(*Call "bds_mem_readBlock" api.*)
///
///bds_mem_readBlock(78,ADR(Readval),100,1);
///
///(*The Readval is to be updated with the asssigned value via the markBlock API*)
///
///
///============================================================================
{attribute 'external_name' := 'cmp_rts_bds_mem_markBlock'}
FUNCTION bds_mem_markBlock : UINT
VAR_INPUT
	///Block number of the NVM Block which marker status has to be changed.
	blockNum_u8: USINT;
	///Data of this variable to be stored in NVM
	dataPtr_u8: POINTER TO USINT;
	///Start address of the NVM sector under the given block number
	startAddress_u16: UINT;
	///Size of the data
	size_u16: UINT;
	///
	///    + TRUE: set the block marker for writing the block during next ECU after run
	///    + FALSE: reset the block marker, means that the block will not be written during next ECU after run
	write_l: BOOL;
END_VAR

END_FUNCTION

// Memory API/NVM/FFI_API/bds_mem_markBlock_ffi
{attribute 'external_name' := 'cmp_rts_bds_mem_markBlock_ffi'}
FUNCTION bds_mem_markBlock_ffi : UINT
VAR_INPUT
	///Block number of the NVM Block which marker status has to be changed.
	blockNum_u8: USINT;
	///Data of this variable to be stored in NVM
	dataPtr_u8: POINTER TO USINT;
	///Start address of the NVM sector under the given block number
	startAddress_u16: UINT;
	///Size of the data
	size_u16: UINT;
	///
	///    + TRUE: set the block marker for writing the block during next ECU after run
	///    + FALSE: reset the block marker, means that the block will not be written during next ECU after run
	write_l: BOOL;
END_VAR

END_FUNCTION

// Memory API/NVM/API/bds_mem_readBlock
///This function copies the data of one NVM block from NVM into respective RAM mirror.
///
///=======
/// Remarks:
///=======
///
///
///    + All RAM mirrors of the application NVM blocks are automatically loaded from system during start up.
///    + This function can be used to restore the RAM mirror of one NVM block with the contents of the NVM during run time.
///    + The |GVL_mem| is given for usage of defines.
///
///----------
/// FFI:
///----------
///    + This API can be used in trusted partitions . For untrusted partitions use |bds_mem_readBlock_ffi|. See Freedom from Interference (FFI) concept for more details.
///    + The blocks which can be read using |bds_mem_readBlock_ffi| are mentioned in page NVM block description.
///
///----------
/// NOTICE:
///----------
///    + This is an asynchronous function. This means that this function already returns as soon as the read request was queued for the NVM server. 
///    + The current read state of a NVM block can be checked with function |bds_mem_getBlockStatus|.
///
///==================================================================		  			===================================================================================================
///Return value    								  									Description
///==================================================================		  			===================================================================================================
///16#0000: BDS_MEM_NO_ERROR_DU16														Reading of block was successfully started.
///16#0001: BDS_MEM_INVALID_BLOCKID_DU16												Invalid Block ID.
///16#0100: BDS_MEM_READBLOCK_ERROR_DU16												Read block could not be started e.g. due to actual block status.
///16#0300: BDS_MEM_READBLOCK_DATASIZE_INVALID_DU16									Read failure as the data size not fitting into NVM Block
///16#0301: BDS_MEM_READBLOCK_DATAPTR_INVALID_DU16										Invalid Data Address
///16#000C: BDS_MEM_FFI_ACCESS_ERROR_DU16												Invalid Access to FFI variant API call.
///
///==================================================================		   			===================================================================================================
///
///
///=======
///Code Example:
///=======
///============================================================================
///
///PROGRAM readPou
///VAR
///
///	ts_mem_read : UINT;
///	
///	Readval: USINT;
///	
///END_VAR
///
///ts_mem_read :=bds_mem_readBlock(78,ADR(Readval),100,1);
///
///  IF(ts_mem_read = 0) THEN
///
///    // read/restore task was successfully started
///  
///  END_IF
///
///============================================================================
{attribute 'external_name' := 'cmp_rts_bds_mem_readBlock'}
FUNCTION bds_mem_readBlock : UINT
VAR_INPUT
	///Block number in which data wanted to be read
	blockNum_u8: USINT;
	///Data of this variable to be read from NVM
	dataPtr_u8: POINTER TO USINT;
	///Start address of the NVM sector under the given block number
	startAddress_u16: UINT;
	///Size of the data
	size_u16: UINT;
END_VAR

END_FUNCTION

// Memory API/NVM/FFI_API/bds_mem_readBlock_ffi
{attribute 'external_name' := 'cmp_rts_bds_mem_readBlock_ffi'}
FUNCTION bds_mem_readBlock_ffi : UINT
VAR_INPUT
	///Block number in which data wanted to be read
	blockNum_u8: USINT;
	///Data of this variable to be read from NVM
	dataPtr_u8: POINTER TO USINT;
	///Start address of the NVM sector under the given block number
	startAddress_u16: UINT;
	///Size of the data
	size_u16: UINT;
END_VAR

END_FUNCTION

// Memory API/NVM/API/bds_mem_getBlockStatus
/// This function gets the current status of one NVM block.
///
///=======
/// Remarks:
///=======
///    + This function must be used to check whether the BSW was successful in loading the NVM blocks during start up.
///    + For more information refer NVM block restoration.
///    + The function can be used to check the result of additional read / write operations which are triggered by the application.
///    + This function can only be used for reading the status of application NVM blocks.
///    + If a NVM block is defined as redundant then a reading error means that none of both NVM blocks could be read successfully.
///    + The |GVL_mem| is given for usage of defines.
///
///----------
/// FFI:
///----------
///This API can be used in trusted partitions . For untrusted partitions use |bds_mem_getBlockStatus_ffi|. See Freedom from Interference (FFI) concept for more details.
///	
///----------
/// NOTICE:
///----------
///
///At the very first startup the NVM blocks will be uninitialized. The BSW will initialize all the data blocks with the value 16#FF.
///
///----------
/// DANGER:
///----------
///
///If the loading of NVM blocks with safety relevant data during start up was not successful then the application must initialize these data with valid values or must enter into a safe state.
///
///==================================================================		  			===================================================================================================
///Return value    								  									Description(Meaning directly after power on)
///==================================================================		  			===================================================================================================
///16#0000: BDS_MEM_NO_ERROR_DU16														Indicates that the previous read operation was completed successfully.
///16#0001: BDS_MEM_INVALID_BLOCKID_DU16												Function bds_mem_getBlockStatus was called with invalid block id.
///16#0300: BDS_MEM_GETBLOCKSTATUS_ERROR_DU16											Function bds_mem_getBlockStatus was not successfully executed.
///16#0301: BDS_MEM_REQ_FAILED_DU16													Indicates that the previous read operation failed.
///16#0302: BDS_MEM_REQ_PENDING_DU16													n.a.
///16#0303: BDS_MEM_REQ_INTEGRITY_FAILED_DU16											Indicates that the previous read operation did not find any valid data for this block on the persistent media. The RAM mirror and NVM block were initialized with 16#FF. The application has to initialize the block with valid data.
///16#0304: BDS_MEM_REQ_BLOCK_SKIPPED_DU16												The NVM block did not yet exist in DFLASH. The RAM mirror and NVM block were initialized with 16#FF. The application has to initialize the block with valid data.
///16#0305: BDS_MEM_REQ_NV_INVALIDATED_DU16											Indicates that the previous read operation only found an invalidated block on the persistent media. The RAM mirror and NVM block were initialized with 16#FF. The application has to initialize the block with valid data.
///16#0308: BDS_MEM_REQ_RESTORED_FROM_ROM_DU16											Indicates that the previous read operation failed e.g., due to CRC failure. Only the RAM mirror was initialized with 16#FF, but the NVM block keeps unchanged. To prevent this error during next read operation the corresponding RAM mirror has to be initialized and written into NVM by the application. 
///16#000C: BDS_MEM_FFI_ACCESS_ERROR_DU16												Invalid Access to FFI variant API call.
///
///==================================================================		   			===================================================================================================
///	
///
///==================================================================		  			===================================================================================================
///Return value    								  									Description(Meaning directly after SW reset)
///==================================================================		  			===================================================================================================
///16#0000: BDS_MEM_NO_ERROR_DU16														Indicates that the previous read operation was completed successfully.
///16#0001: BDS_MEM_INVALID_BLOCKID_DU16												Function bds_mem_getBlockStatus was called with invalid block id.
///16#0300: BDS_MEM_GETBLOCKSTATUS_ERROR_DU16											Function bds_mem_getBlockStatus was not successfully executed.
///16#0301: BDS_MEM_REQ_FAILED_DU16													Indicates that the previous read operation failed.
///16#0302: BDS_MEM_REQ_PENDING_DU16													n.a.
///16#0303: BDS_MEM_REQ_INTEGRITY_FAILED_DU16											Indicates that the previous read operation did not find any valid data for this block on the persistent media. The RAM mirror and NVM block were initialized with 16#FF. The application has to initialize the block with valid data.
///16#0304: BDS_MEM_REQ_BLOCK_SKIPPED_DU16												n.a.
///16#0305: BDS_MEM_REQ_NV_INVALIDATED_DU16											Indicates that the previous read operation only found an invalidated block on the persistent media. The RAM mirror and NVM block were initialized with 16#FF. The application has to initialize the block with valid data.
///16#0308: BDS_MEM_REQ_RESTORED_FROM_ROM_DU16											Indicates that the previous read operation failed e.g., due to CRC failure. Only the RAM mirror was initialized with 16#FF, but the NVM block keeps unchanged. To prevent this error during next read operation the corresponding RAM mirror has to be initialized and written into NVM by the application. 
///16#000C: BDS_MEM_FFI_ACCESS_ERROR_DU16												Invalid Access to FFI variant API call.
///
///==================================================================		   			===================================================================================================
///	
///
///==================================================================		  			===================================================================================================
///Return value    								  									Description(Meaning after |bds_mem_readBlock|)
///==================================================================		  			===================================================================================================
///16#0000: BDS_MEM_NO_ERROR_DU16														Indicates that the previous read operation was completed successfully.
///16#0001: BDS_MEM_INVALID_BLOCKID_DU16												Function bds_mem_getBlockStatus was called with invalid block id.
///16#0300: BDS_MEM_GETBLOCKSTATUS_ERROR_DU16											Function bds_mem_getBlockStatus was not successfully executed.
///16#0301: BDS_MEM_REQ_FAILED_DU16													Indicates that the previous read operation failed.
///16#0302: BDS_MEM_REQ_PENDING_DU16													Indicates that the previous read operation is still ongoing.
///16#0303: BDS_MEM_REQ_INTEGRITY_FAILED_DU16											Indicates that the previous read operation did not find any valid data for this block on the persistent media. The RAM mirror and NVM block were initialized with 16#FF. The application has to initialize the block with valid data.
///16#0304: BDS_MEM_REQ_BLOCK_SKIPPED_DU16												n.a.
///16#0305: BDS_MEM_REQ_NV_INVALIDATED_DU16											Indicates that the previous read operation only found an invalidated block on the persistent media. The RAM mirror and NVM block were initialized with 16#FF. The application has to initialize the block with valid data.
///16#0308: BDS_MEM_REQ_RESTORED_FROM_ROM_DU16											Indicates that the previous read operation failed e.g., due to CRC failure. Only the RAM mirror was initialized with 16#FF, but the NVM block keeps unchanged. To prevent this error during next read operation the corresponding RAM mirror has to be initialized and written into NVM by the application. 
///16#000C: BDS_MEM_FFI_ACCESS_ERROR_DU16												Invalid Access to FFI variant API call.
///
///==================================================================		   			===================================================================================================
///	
///
///==================================================================		  			===================================================================================================
///Return value    								  									Description(Meaning after |bds_mem_writeBlock|)
///==================================================================		  			===================================================================================================
///16#0000: BDS_MEM_NO_ERROR_DU16														Indicates that the previous write operation was completed successfully
///16#0001: BDS_MEM_INVALID_BLOCKID_DU16												Function bds_mem_getBlockStatus was called with invalid block id.
///16#0300: BDS_MEM_GETBLOCKSTATUS_ERROR_DU16											Function bds_mem_getBlockStatus was not successfully executed.
///16#0301: BDS_MEM_REQ_FAILED_DU16													Indicates that the previous write operation failed.
///16#0302: BDS_MEM_REQ_PENDING_DU16													Indicates that the previous write operation is still ongoing.
///16#0303: BDS_MEM_REQ_INTEGRITY_FAILED_DU16											n.a.
///16#0304: BDS_MEM_REQ_BLOCK_SKIPPED_DU16												n.a.
///16#0305: BDS_MEM_REQ_NV_INVALIDATED_DU16											n.a.
///16#0308: BDS_MEM_REQ_RESTORED_FROM_ROM_DU16											n.a.
///16#000C: BDS_MEM_FFI_ACCESS_ERROR_DU16												Invalid Access to FFI variant API call.
///
///==================================================================		   			===================================================================================================
///
///=======
///Code Example:
///=======
///============================================================================
///
///PROGRAM nvm
///
///VAR
///
///	status_u16: uint;	
///	
///END_VAR
///
///status_u16:=bds_mem_getBlockStatus(bds_mem_nvmBlock03_512_R_D);
///
///(*evaluate the status of NVM block 3*)
///
///if (BDS_MEM_NO_ERROR_DU16 = status_u16) THEN
///
///	(*last read/write operation was completed successfully*)
///
///END_IF
///
///============================================================================
///
///	
{attribute 'external_name' := 'cmp_rts_bds_mem_getBlockStatus'}
FUNCTION bds_mem_getBlockStatus : UINT
VAR_INPUT
	///Block id of the NVM block which is to be checked. The list of available block ids is available in NVM Block Description. 
	blockId_u16: UINT;
END_VAR

END_FUNCTION

// Memory API/NVM/FFI_API/bds_mem_getBlockStatus_ffi
{attribute 'external_name' := 'cmp_rts_bds_mem_getBlockStatus_ffi'}
FUNCTION bds_mem_getBlockStatus_ffi : UINT
VAR_INPUT
	///Block id of the NVM block which is to be checked. The list of available block ids is available in NVM Block Description. 
	blockId_u16: UINT;
END_VAR

END_FUNCTION

// Memory API/NVM/API/bds_mem_writeBlock
/// This function writes the data from the variable(s) of the RAM mirror into corresponding NVM block.
///
///=======
/// Remarks:
///=======
///
///    + This function can be used to store the RAM mirror already before execution of after run.
///    + All RAM mirrors of the application NVM blocks which have been marked previously with function |bds_mem_markBlock| are automatically stored to NVM during after run.
///    + The |GVL_mem| is given for usage of defines.
///
///----------
/// FFI:
///----------
///    + This API can be used in trusted partitions . For untrusted partitions use |bds_mem_writeBlock_ffi|. See Freedom from Interference (FFI) concept for more details.
///    + The blocks which can be written using |bds_mem_writeBlock_ffi| are mentioned in page NVM block description.
///
///----------
/// NOTICE:
///----------
///    + This is an asynchronous function. This means that this function already returns as soon as the write request was queued for the NVM server. 
///    + The current write state of a NVM block can be checked with function |bds_mem_getBlockStatus|.
///
///----------
/// CAUTION:
///----------
///    + Do not use this function with high frequency in cyclic tasks because the DFlash cells of the NVM have limited number of write cycles! 
///    + This function writes the data physically into the DFlash even so if the data was not changed!
///    + Do not call this function more often than really required or use the function bds_mem_markBlock for a single storage process during after run.
///
///==================================================================		  			===================================================================================================
///Return value    								  									Description
///==================================================================		  			===================================================================================================
///16#0000: BDS_MEM_NO_ERROR_DU16														Writing of block was successfully started.
///16#0001: BDS_MEM_INVALID_BLOCKID_DU16												Invalid Block ID.
///16#0200: BDS_MEM_WRITEBLOCK_ERROR_DU16												Write block could not be started e.g., due to actual block status
///16#0300: BDS_MEM_WRITEBLOCK_DATASIZE_INVALID_DU16									Write failure as the data size not fitting into NVM Block
///16#0301: BDS_MEM_WRITEBLOCK_DATAPTR_INVALID_DU16									Invalid Data Address
///16#000C: BDS_MEM_FFI_ACCESS_ERROR_DU16												Invalid Access to FFI variant API call.
///
///==================================================================		   			===================================================================================================
///
///
///=======
///Code Example:
///=======
///============================================================================
///
///PROGRAM writePou
///VAR
///
///	Writeval_u8:USINT:=0;
///	
///	ts_mem_write : UINT;
///	
///	flagWrite: USINT:=0;
///	
///	Readval_u8: USINT:=0;
///	
///END_VAR
///	
///END_IF
///
///IF(flagWrite=0) THEN
///
///	ts_mem_write:=bds_mem_writeBlock(78,ADR(Writeval_u8),100,1);
///	
///	flagWrite:=1;
///	
///	IF(ts_mem_write = 0) THEN
///
///    // write task was successfully started  
///	
/// END_IF
///	
///END_IF
///
/// (*The readBlock data pointer should be updated with data written in the respective block*)
///
///bds_mem_readBlock(78,ADR(Readval_u8),100,1);
///
///
///============================================================================
{attribute 'external_name' := 'cmp_rts_bds_mem_writeBlock'}
FUNCTION bds_mem_writeBlock : UINT
VAR_INPUT
	///Block number in which data has to be written
	blockNum_u8: USINT;
	///Data of this variable to be stored in NVM
	dataPtr_u8: POINTER TO USINT;
	///Start address of the NVM sector under the given block number
	startAddress_u16: UINT;
	///Size of the data
	size_u16: UINT;
END_VAR

END_FUNCTION

// Memory API/NVM/FFI_API/bds_mem_writeBlock_ffi
{attribute 'external_name' := 'cmp_rts_bds_mem_writeBlock_ffi'}
FUNCTION bds_mem_writeBlock_ffi : UINT
VAR_INPUT
	///Block number in which data has to be written
	blockNum_u8: USINT;
	///Data of this variable to be stored in NVM
	dataPtr_u8: POINTER TO USINT;
	///Start address of the NVM sector under the given block number
	startAddress_u16: UINT;
	///Size of the data
	size_u16: UINT;
END_VAR

END_FUNCTION

// System API/SYS/API/bds_sys_resetINH
///This function sets the Inhibit signal to reset.
///=======
/// Remarks:
///=======
///    + With the activation of signals Inhibit1 or Inhibit2 the power output stages are disabled.
///    + After reactivation of the signals this function has to be called to enable the inhibit hardware again.
///    + Restart of signal INH allowed if previous reset is finished. 
///    + The |GVL_sys| is given for usage of defines.
///
///----------
/// FFI:
///----------
///This API can be used in trusted partitions only. See Freedom from Interference (FFI) concept for more details.
///
///---------
///  CAUTION:
///---------
///This reset happens as a background task. So, it needs maximum 3ms to reset the inhibit signal.
///	
///==================================================================		  			===================================================================================================
///Return value    								  									Description
///==================================================================		  			===================================================================================================
///None																				None
///
///==================================================================		   			===================================================================================================
///
///=======
///Code Example:
///=======
///============================================================================
///
///PROGRAM appl_10ms_task
///
///VAR
///
///END_VAR
///
///(* reset signal INH after a activation of inhibit *)
///
///bds_sys_resetINH();
///
///
///============================================================================
///
{attribute 'external_name' := 'cmp_rts_bds_sys_resetINH'}
FUNCTION bds_sys_resetINH : BOOL

END_FUNCTION

// System API/SYS/API/bds_sys_setVSS
///This function sets the sensor supply voltage to the given state.
///=======
/// Remarks:
///=======
///    + After startup of the ECU all VSS are enabled. 
///    + For the further information regarding the recovery of the sensor supplies after short circuits see Cyclic monitoring checks.
///    + The |GVL_sys| is given for usage of defines.
///    + Import the bds_rts_ec.xml to use the enums. (Refer example below).
///	
///----------
/// FFI:
///----------
///This API can be used in trusted partitions only. See Freedom from Interference (FFI) concept for more details.
///
///==================================================================		  			===================================================================================================
///Return value    								  									Description
///==================================================================		  			===================================================================================================
///16#00																				No error.
///16#01																				A parameter is invalid.
///16#02																				Function call was erroneous.
///
///==================================================================		   			===================================================================================================
///
///=======
///Code Example:
///=======
///============================================================================
///
///PROGRAM PLC_PRG
///
///  VAR
///
///  END_VAR
///
///(* switch VSS1 on *)
///
///bds_sys_setVSS(bds_sys_vss_signal_te.VSS1, STD_ON);
///
///============================================================================
///
{attribute 'external_name' := 'cmp_rts_bds_sys_setVSS'}
FUNCTION bds_sys_setVSS : USINT
VAR_INPUT
	///The assigned signal name.
	signal_e: UINT;
	///States of the sensor supply.
	///    + STD_OFF  - Disable the VSS,
	///    + STD_ON   -  Enable the VSS (default).
	state_u8: USINT;
END_VAR

END_FUNCTION

// System API/SYS/API/bds_sys_startLoader
///This function starts the program loader.
///=======
/// Remarks:
///=======
///    + This function should be called to flash the ECU.
///    + Before this function call bds_sys_startLoader(), the memory blocks ,which need to be saved into NVM (NVM general description), should be marked by calling the  function |bds_mem_markBlock|. Thus, during reset preparation marked memory block is saved into NVM and it can be retrieved after reset.
///    + The |GVL_sys| is given for usage of defines.
///
///	
///----------
/// FFI:
///----------
///This API can be used in trusted partitions only. See Freedom from Interference (FFI) concept for more details.
///
///==================================================================		  			===================================================================================================
///Return value    								  									Description
///==================================================================		  			===================================================================================================
///None																				None
///
///==================================================================		   			===================================================================================================
///
///=======
///Code Example:
///=======
///============================================================================
///
///PROGRAM appl_1ms_task
///
///VAR
///
///    Mark_writeval: USINT:=0;
///
///END_VAR
///
///(*Call the markblock API. Mark the block(eg:3rd block) which has to be written during afterrun cycle in either cyclic task or calling once & assign a value to Mark_writeval*)
///
///bds_mem_markBlock(3,ADR(Mark_writeval),1,1,TRUE);
///
///bds_sys_startLoader(TRUE, 0x1234);
///
///============================================================================
///
{attribute 'external_name' := 'cmp_rts_bds_sys_startLoader'}
FUNCTION bds_sys_startLoader : BOOL
VAR_INPUT
	///If the “NVMWrite_l” flag is set to the following values the behaviour is different,
	///TRUE   : It starts the loader after the queue of NVM is empty.
	///FALSE  : It starts the loader directly.
	NVMWrite_l: BOOL;
	///User-defined value can be used for application purpose in CB.
	userData_u32: UDINT;
END_VAR

END_FUNCTION

// Diagnostics API/UDS/API/bds_uds_disable
///This function is to disable/enable the BSW UDS stack
///
///=======
/// Remarks:
///=======
///    + By default the UDS stack is enabled by the BSW.
///    + The |GVL_uds| is given for usage of defines.
///
///----------
/// FFI:
///----------
///This API can be used in trusted partitions only. See Freedom from Interference (FFI) concept for more details.
///
///==================================================================		  			===================================================================================================
///Return value    								  									Description
///==================================================================		  			===================================================================================================
///None.																				-
///
///==================================================================		   			===================================================================================================
///=======
///Code Example:
///=======
///============================================================================
///
///PROGRAM PLC_PRG
///  VAR
///	FLAG:BOOL;
/// END_VAR
///  
///IF FLAG:=False THEN
///
///	(*disable the UDS stack*)
///	
///	bds_uds_disable(TRUE); 
///
///	FLAG:= TRUE;
///
///END_IF
///
///============================================================================
{attribute 'external_name' := 'cmp_rts_bds_uds_disable'}
FUNCTION bds_uds_disable : BOOL
VAR_INPUT
	///The parameter defines
	///    + TRUE - UDS stack is disabled
	///    + FALSE - UDS stack is enabled
	uds_disableFlg_l: BOOL;
END_VAR

END_FUNCTION

// Diagnostics API/UDS/API/bds_uds_GetActiveDid
///This function gets the active DID from Diagnostics Communication.
///
///=======
/// Remarks:
///=======
///    + Data identifiers can be added from easyConfig with the specified ranges.
///    + Access levels of security and session can be mapped from easyConfig.
///    + |bds_sys_memByteCopy| API to be used to fill the data into buffer.
///    + The |GVL_uds| is given for usage of defines.
///
///----------
/// FFI:
///----------
///This API can be used in trusted partitions only. See Freedom from Interference (FFI) concept for more details.
///
///==================================================================		  			===================================================================================================
///Return value    								  									Description
///==================================================================		  			===================================================================================================
///0																					Valid Data Identifier
///1																					Invalid Data Identifier
///
///==================================================================		   			===================================================================================================
///=======
///Code Example:
///=======
///============================================================================
///
///FUNCTION POU_1 : BYTE
///VAR_INPUT
///
///    can_data : POINTER TO BYTE;
///END_VAR
///
///
///bds_uds_GetActiveDid(ADR(DidValue_u16));
///
///IF (DidValue_u16=16#100)
///
///  THEN bds_uds_setCallbackStatus(0);(*positive response for DID 16#100*)
///  
///END_IF
///
///
///(*Registering callback*)
///
///PROGRAM POU_10
///VAR
///
///	flag_1 : BOOL := 1; 
///
///END_VAR
///
///IF ( flag_1)
///
///    THEN bds_uds_registerDidReadCallback (ADR(POU_1));
///
///    flag_1 := 0;(*To make api call once in application*)
///
///END_IF
///
///============================================================================
{attribute 'external_name' := 'cmp_rts_bds_uds_GetActiveDid'}
FUNCTION bds_uds_GetActiveDid : USINT
VAR_INPUT
	///Reference of variable where the active DataIdentifier will be saved by the API. 
	Get_DID_u16: POINTER TO UINT;
END_VAR

END_FUNCTION

// Diagnostics API/UDS/API/bds_uds_setCallbackStatus
///This function will set the return value for the UDS DID & Routine Control callbacks used in the UDS module.
///
///=======
/// Remarks:
///=======
///    + This is the mandatory API to be used to set the callback status.
///    + The |GVL_uds| is given for usage of defines.
///
///----------
/// FFI:
///----------
///This API can be used in trusted partitions only. See Freedom from Interference (FFI) concept for more details.
///
///==================================================================		  			===================================================================================================
///Return value    								  									Description
///==================================================================		  			===================================================================================================
///0																					No error
///1																					Invalid pointer
///
///==================================================================		   			===================================================================================================
///
///=======
///Code Example:
///=======
///============================================================================
///
///FUNCTION POU_1 : BYTE
///VAR_INPUT
///
///    can_data : POINTER TO BYTE;
///END_VAR
///
///VAR
///    data_au8 : ARRAY[0..8] OF BYTE;
///	
///    i1: BYTE;
///	
///    DidValue_u16: UINT;
///	
///    set_u8: USINT;
///END_VAR
///
///
///bds_uds_GetActiveDid(ADR(DidValue_u16));
///
///IF (DidValue_u16=16#100)
///
///  THEN bds_uds_setCallbackStatus(0);(*positive response for DID 16#100*)
///  
///END_IF
///
///IF (DidValue_u16=16#200) 
///
///  THEN  bds_uds_setCallbackStatus(1);(*negative response for DID 16#200*)
///  
///END_IF
///
///FOR i1 := 0 TO 8 BY 1 DO
///can_data[i1]  := data_au8[i1];
///END_FOR;
///POU_1 :=1;
///
///(*Registering callback*)
///
///PROGRAM POU_10
///VAR
///
///	flag_1 : BOOL := 1;
///	
///    flag_2 : BOOL := 1; 
///   
///    flag_3 : BOOL := 1;    
///
///END_VAR
///
///IF ( flag_1)
///
///    THEN bds_uds_registerDidReadCallback (ADR(POU_1));
///
///    flag_1 := 0;
///
///END_IF
///
///IF ( flag_2)
///
///    THEN bds_uds_registerDidWriteCallback (ADR(POU_2));
///
///    flag_2 := 0;
///
///END_IF
///
///IF ( flag_3)
///
///    THEN bds_uds_registerRoutineF000Callback (ADR(POU_3));
///
///    flag_3 := 0;
///
///END_IF
///
///
///============================================================================
{attribute 'external_name' := 'cmp_rts_bds_uds_setCallbackStatus'}
FUNCTION bds_uds_setCallbackStatus : BOOL
VAR_INPUT
	/// 
	///possible vales:
	///   + E_OK(0): Positive response
	///   + E_NOT_OK(1) : negative response
	///   + Request Pending(0x0010): This asynchronous function was not yet completed and must be called again with the same parameter values.
	status_u8: USINT;
END_VAR

END_FUNCTION

// Diagnostics API/UDS/API/bds_uds_registerDidReadCallback
///This function registers the callback for DID read operation.
///
///=======
/// Remarks:
///=======
///    + This is the mandatory API to be used if the DID parameter/ process data need to be read.
///    + The |GVL_uds| is given for usage of defines.
///
///----------
/// FFI:
///----------
///This API can be used in trusted partitions only. See Freedom from Interference (FFI) concept for more details.
///
///==================================================================		  			===================================================================================================
///Return value    								  									Description
///==================================================================		  			===================================================================================================
///0																					No error
///1																					Invalid pointer
///
///==================================================================		   			===================================================================================================
///
///=======
///Code Example:
///=======
///============================================================================
///
///FUNCTION POU_1 : BYTE
///VAR_INPUT
///
///    can_data : POINTER TO BYTE;
///END_VAR
///
///VAR
///    data_au8 : ARRAY[0..8] OF BYTE;
///	
///    i1: BYTE;
///	
///    DidValue_u16: UINT;
///	
///    set_u8: USINT;
///END_VAR
///
///
///bds_uds_GetActiveDid(ADR(DidValue_u16));
///
///IF (DidValue_u16=16#100)
///
///  THEN bds_uds_setCallbackStatus(0);(*positive response for DID 16#100*)
///  
///END_IF
///
///IF (DidValue_u16=16#200) 
///
///  THEN  bds_uds_setCallbackStatus(1);(*negative response for DID 16#200*)
///  
///END_IF
///
///FOR i1 := 0 TO 8 BY 1 DO
///can_data[i1]  := data_au8[i1];
///END_FOR;
///POU_1 :=1;
///
///(*Registering callback*)
///
///PROGRAM POU_10
///VAR
///
///	flag_1 : BOOL := 1;
///	
///    flag_2 : BOOL := 1; 
///   
///    flag_3 : BOOL := 1;    
///
///END_VAR
///
///IF ( flag_1)
///
///    THEN bds_uds_registerDidReadCallback (ADR(POU_1));
///
///    flag_1 := 0;(*To make api call once in application*)
///
///END_IF
///
///IF ( flag_2)
///
///    THEN bds_uds_registerDidWriteCallback (ADR(POU_1));
///
///    flag_2 := 0;(*To make api call once in application*)
///
///END_IF
///
///IF ( flag_3)
///
///    THEN bds_uds_registerRoutineF000Callback (ADR(POU_3));
///
///    flag_3 := 0;(*To make api call once in application*)
///
///END_IF
///
///
///============================================================================
{attribute 'external_name' := 'cmp_rts_bds_uds_registerDidReadCallback'}
FUNCTION bds_uds_registerDidReadCallback : USINT
VAR_INPUT
	///Function pointer with argument of UINT8 data pointer
	func_pf: POINTER TO BOOL;
END_VAR

END_FUNCTION

